TYPE U_APP_STATE :
UNION
  stState             : ST_TOWER_STATE;
  byState   AT %i*    : ARRAY[1..SIZEOF(ST_TOWER_STATE)] OF BYTE;
END_UNION
END_TYPE

(* stored: Version 1.1.0.1
   DUT U_APP_STATE: Id {77441d2c-f847-4ff3-a6c9-65b646e727c3} *)
